(* Logix 5000 project; controller SigmaAldrich vendor 1 type 14 code 77 rev 15.4; software revision 15.02; part 3 of 3 *)
(* tags used below, declared in another part *)
   Airlock_N1068_E_Stop_OSR : BOOL;
   Airlock_N1068_Violation_MDI_Bit : BOOL;
   Airlock_N1068_Violation_MDI_OSR : BOOL;
   Annuciator_Bit_Airlock_N1068 : BOOL;
   Door_N1068A_Timer : TIMER;
   Door_N1068B_Timer : TIMER;
   MDI_Violation_N1068_Bit : BOOL;
   N1068_Airlock_Latch : BOOL;
   N1068_Emergency_Release_Latch : BOOL;
   N1068B_Door_Latch_Bit : BOOL;
(* MainProgram, continued *)

ROUTINE DI15_N1068   (* ladder *)
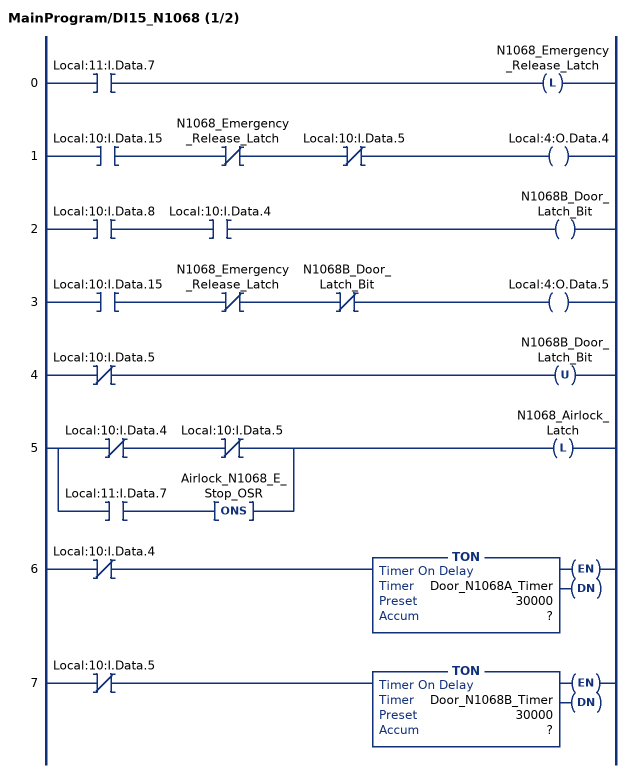
   0: XIC(Local:11:I.Data.7)OTL(N1068_Emergency_Release_Latch);
   1: XIC(Local:10:I.Data.15)XIO(N1068_Emergency_Release_Latch)XIO(Local:10:I.Data.5)OTE(Local:4:O.Data.4);
   2: XIC(Local:10:I.Data.8)XIC(Local:10:I.Data.4)OTE(N1068B_Door_Latch_Bit);
   3: XIC(Local:10:I.Data.15)XIO(N1068_Emergency_Release_Latch)XIO(N1068B_Door_Latch_Bit)OTE(Local:4:O.Data.5);
   4: XIO(Local:10:I.Data.5)OTU(N1068B_Door_Latch_Bit);
   5: [XIO(Local:10:I.Data.4) XIO(Local:10:I.Data.5) ,XIC(Local:11:I.Data.7) ONS(Airlock_N1068_E_Stop_OSR) ]OTL(N1068_Airlock_Latch);
   6: XIO(Local:10:I.Data.4)TON(Door_N1068A_Timer,?,?);
   7: XIO(Local:10:I.Data.5)TON(Door_N1068B_Timer,?,?);
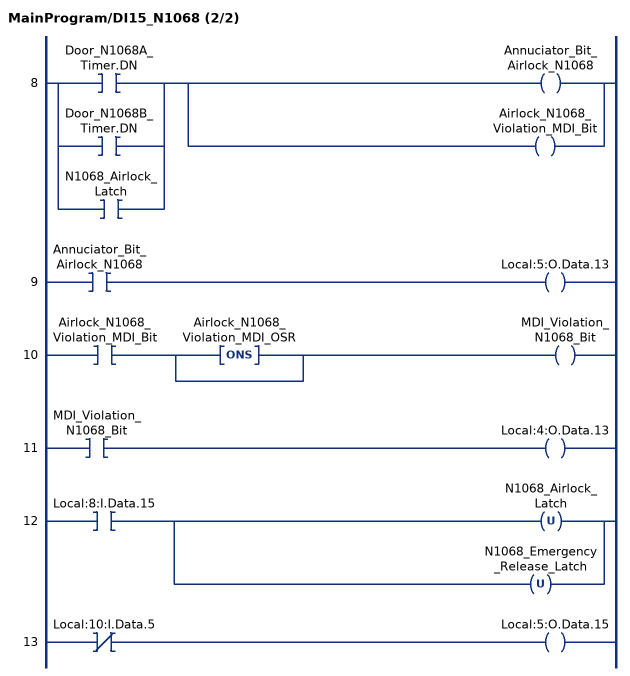
   8: [XIC(Door_N1068A_Timer.DN) ,XIC(Door_N1068B_Timer.DN) ,XIC(N1068_Airlock_Latch) ][OTE(Annuciator_Bit_Airlock_N1068) ,OTE(Airlock_N1068_Violation_MDI_Bit) ];
   9: XIC(Annuciator_Bit_Airlock_N1068)OTE(Local:5:O.Data.13);
   10: XIC(Airlock_N1068_Violation_MDI_Bit)[ONS(Airlock_N1068_Violation_MDI_OSR) ,]OTE(MDI_Violation_N1068_Bit);
   11: XIC(MDI_Violation_N1068_Bit)OTE(Local:4:O.Data.13);
   12: XIC(Local:8:I.Data.15)[OTU(N1068_Airlock_Latch) ,OTU(N1068_Emergency_Release_Latch) ];
   13: XIO(Local:10:I.Data.5)OTE(Local:5:O.Data.15);
END_ROUTINE

ROUTINE Door_N1137A   (* ladder *)
END_ROUTINE

ROUTINE Doors_N1034A_34B_37B   (* ladder *)
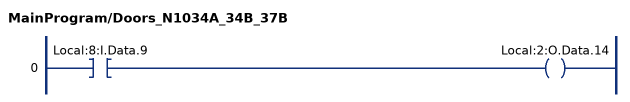
   0: XIC(Local:8:I.Data.9)OTE(Local:2:O.Data.14);
END_ROUTINE

ROUTINE MainRoutine   (* ladder *)
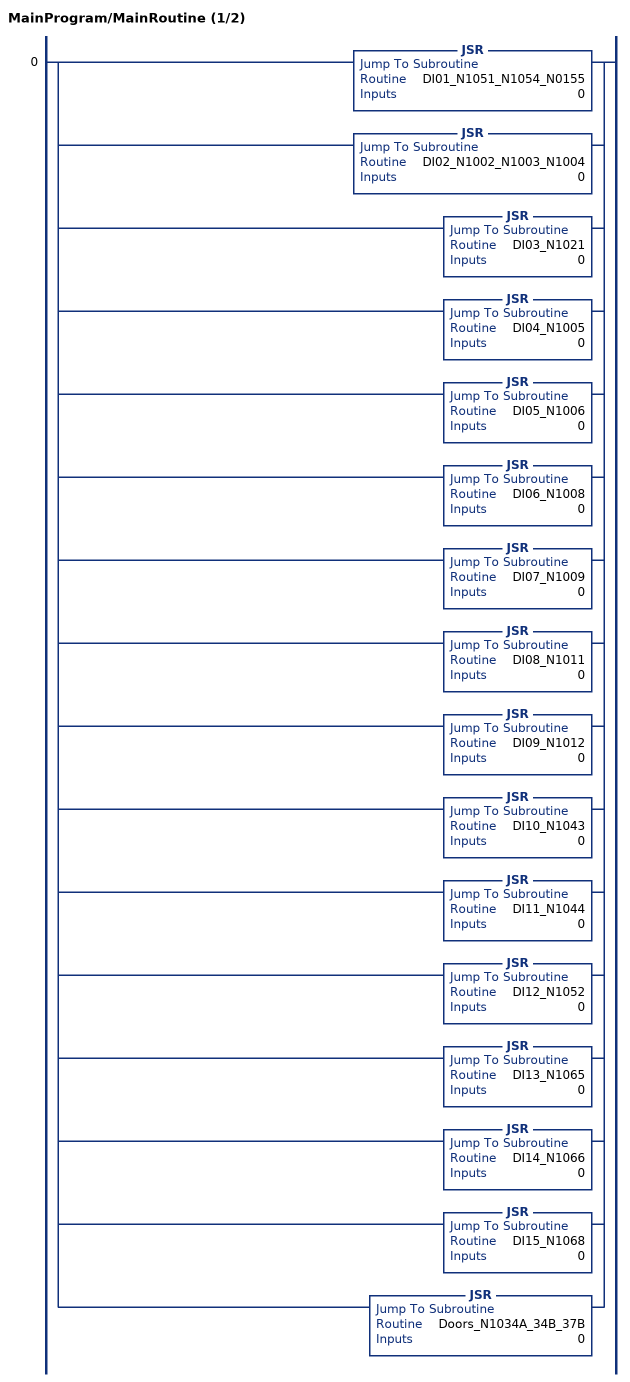
   0: [JSR(DI01_N1051_N1054_N0155,0) ,JSR(DI02_N1002_N1003_N1004,0) ,JSR(DI03_N1021,0) ,JSR(DI04_N1005,0) ,JSR(DI05_N1006,0) ,JSR(DI06_N1008,0) ,JSR(DI07_N1009,0) ,JSR(DI08_N1011,0) ,JSR(DI09_N1012,0) ,JSR(DI10_N1043,0) ,JSR(DI11_N1044,0) ,JSR(DI12_N1052,0) ,JSR(DI13_N1065,0) ,JSR(DI14_N1066,0) ,JSR(DI15_N1068,0) ,JSR(Doors_N1034A_34B_37B,0) ];
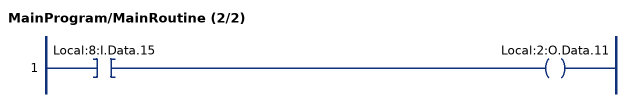
   1: XIC(Local:8:I.Data.15)OTE(Local:2:O.Data.11);
END_ROUTINE
END_PROGRAM
